// TIA Portal V14 SP1 export
// export: Created 2000-01-01T00:00:00.0000000Z, ExportSetting WithDefaults, WithReadOnly
DATA_BLOCK "MCP_RC_DB"   // DB9801
{ S7_Optimized_Access := 'FALSE' }
   VAR
      Count : Int := 3;
      Motor : "MCP_RC_UDT";
   END_VAR
BEGIN
END_DATA_BLOCK
